        string sColour
    utBorder Border
      [0]
        num nBorderWidth
        string sBorderColour
        string sBorderStyle
    utCommon Common
      [0]
        string sID = "lbl_Title"
        string sPage = "Disk://SmartTCP_CS9/ts2/interface/Page_Main"
        string sText = "史陶比尔工具标定 - SmartTCP"
    utData Data
      [0]
        bool bStatus
        num nVal = 99
    utEvents Events
      [0]
        bool bClick
        bool bMouseDown
        bool bMouseUp
    utText Text
      [0]
        num nFontSize
        string sFontFamily
        string sFontStyle
        string sFontWeight
        string sTextAlignment
public utLabel utLbl_Tool
  [0]
    utAppearance Appearance
      [0]
        bool bVisibility
        string sBackgroundColour = "#FFFFFF"
        string sColour
    utBorder Border
      [0]
        num nBorderWidth
        string sBorderColour
        string sBorderStyle
    utCommon Common
      [0]
        string sID = "lbl_Tool"
        string sPage = "Disk://SmartTCP_CS9/ts2/interface/Page_Main"
        string sText = "工具："
    utData Data
      [0]
        bool bStatus
        num nVal = 99
    utEvents Events
      [0]
        bool bClick
        bool bMouseDown
        bool bMouseUp
    utText Text
      [0]
        num nFontSize
        string sFontFamily
        string sFontStyle
        string sFontWeight
        string sTextAlignment
public utLabel utLbl_ToolValue_Data[6]
  [0]
    utAppearance Appearance
      [0]
        bool bVisibility
        string sBackgroundColour = "#FFFFFF"
        string sColour
    utBorder Border
      [0]
        num nBorderWidth
        string sBorderColour
        string sBorderStyle
    utCommon Common
      [0]
        string sID = "utLbl_ToolValue_Data0"
        string sPage = "Disk://SmartTCP_CS9/ts2/interface/Page_Container_Test"
        string sText = "120    "
    utData Data
      [0]
        bool bStatus
        num nVal = 99
    utEvents Events
      [0]
        bool bClick
        bool bMouseDown
        bool bMouseUp
    utText Text
      [0]
        num nFontSize
        string sFontFamily
        string sFontStyle
        string sFontWeight
        string sTextAlignment
  [1]
    utAppearance Appearance
      [0]
        bool bVisibility
        string sBackgroundColour = "#FFFFFF"
        string sColour
    utBorder Border
      [0]
        num nBorderWidth
        string sBorderColour
        string sBorderStyle
    utCommon Common
      [0]
        string sID = "utLbl_ToolValue_Data1"
        string sPage = "Disk://SmartTCP_CS9/ts2/interface/Page_Container_Test"
        string sText = "55    "
    utData Data
      [0]
        bool bStatus
        num nVal = 99
    utEvents Events
      [0]
        bool bClick
        bool bMouseDown
        bool bMouseUp
    utText Text
      [0]
        num nFontSize
        string sFontFamily
        string sFontStyle
        string sFontWeight
        string sTextAlignment
  [2]
    utAppearance Appearance
      [0]
        bool bVisibility
        string sBackgroundColour = "#FFFFFF"
        string sColour
    utBorder Border
      [0]
        num nBorderWidth
        string sBorderColour
        string sBorderStyle
    utCommon Common
      [0]
        string sID = "utLbl_ToolValue_Data2"
        string sPage = "Disk://SmartTCP_CS9/ts2/interface/Page_Container_Test"
        string sText = "0    "
    utData Data
      [0]
        bool bStatus
        num nVal = 99
    utEvents Events
      [0]
        bool bClick
        bool bMouseDown
        bool bMouseUp
    utText Text
      [0]
        num nFontSize
        string sFontFamily
        string sFontStyle
        string sFontWeight
        string sTextAlignment
  [3]
    utAppearance Appearance
      [0]
        bool bVisibility
        string sBackgroundColour = "#FFFFFF"
        string sColour
    utBorder Border
      [0]
        num nBorderWidth
        string sBorderColour
        string sBorderStyle
    utCommon Common
      [0]
        string sID = "utLbl_ToolValue_Data3"
        string sPage = "Disk://SmartTCP_CS9/ts2/interface/Page_Container_Test"
        string sText = "0    "
    utData Data
      [0]
        bool bStatus
        num nVal = 99
    utEvents Events
      [0]
        bool bClick
        bool bMouseDown
        bool bMouseUp
    utText Text
      [0]
        num nFontSize
        string sFontFamily
        string sFontStyle
        string sFontWeight
        string sTextAlignment
  [4]
    utAppearance Appearance
      [0]
        bool bVisibility
        string sBackgroundColour = "#FFFFFF"
        string sColour
    utBorder Border
      [0]
        num nBorderWidth
        string sBorderColour
        string sBorderStyle
    utCommon Common
      [0]
        string sID = "utLbl_ToolValue_Data4"
        string sPage = "Disk://SmartTCP_CS9/ts2/interface/Page_Container_Test"
        string sText = "0    "
    utData Data
      [0]
        bool bStatus
        num nVal = 99
    utEvents Events
      [0]
        bool bClick
        bool bMouseDown
        bool bMouseUp
    utText Text
      [0]
        num nFontSize
        string sFontFamily
        string sFontStyle
        string sFontWeight
        string sTextAlignment
  [5]
    utAppearance Appearance
      [0]
        bool bVisibility
        string sBackgroundColour = "#FFFFFF"
        string sColour
    utBorder Border
      [0]
        num nBorderWidth
        string sBorderColour
        string sBorderStyle
    utCommon Common
      [0]
        string sID = "utLbl_ToolValue_Data5"
        string sPage = "Disk://SmartTCP_CS9/ts2/interface/Page_Container_Test"
        string sText = "0    "
    utData Data
      [0]
        bool bStatus
        num nVal = 99
    utEvents Events
      [0]
        bool bClick
        bool bMouseDown
        bool bMouseUp
    utText Text
      [0]
        num nFontSize
        string sFontFamily
        string sFontStyle
        string sFontWeight
        string sTextAlignment
public utLabel utLbl_Tool_Data
  [0]
    utAppearance Appearance
      [0]
        bool bVisibility
        string sBackgroundColour = "#FFFFFF"
        string sColour
    utBorder Border
      [0]
        num nBorderWidth
        string sBorderColour
        string sBorderStyle
    utCommon Common
      [0]
        string sID = "lbl_Tool_Data"
        string sPage = "Disk://SmartTCP_CS9/ts2/interface/Page_Main"
        string sText = "tFlange"
    utData Data
      [0]
        bool bStatus
        num nVal = 99
    utEvents Events
      [0]
        bool bClick
        bool bMouseDown
        bool bMouseUp
    utText Text
      [0]
        num nFontSize
        string sFontFamily
        string sFontStyle
        string sFontWeight
        string sTextAlignment
public utText utTxt_OffsetValue_Data[6]
  [0]
    utAppearance Appearance
      [0]
        bool bVisibility
        string sBackgroundColour = "#EEFF00"
        string sColour
    utBorder Border
      [0]
        string sBorderColour
        string sBorderSytle
        string sBorderWidth
    utCommon Common
      [0]
        bool bDisabled
        num nValue
        string sID = "utTxt_OffsetValue_Data0"
        string sPage = "Disk://SmartTCP_CS9/ts2/interface/Page_Container_Test"
        string sValue
    utText Text
      [0]
        num nFontSize
        string sFontFamily
        string sFontStyle
        string sFontWeight
        string sTextAlignment
  [1]
    utAppearance Appearance
      [0]
        bool bVisibility
        string sBackgroundColour = "#EEFF00"
        string sColour
    utBorder Border
      [0]
        string sBorderColour
        string sBorderSytle
        string sBorderWidth
    utCommon Common
      [0]
        bool bDisabled
        num nValue
        string sID = "utTxt_OffsetValue_Data1"
        string sPage = "Disk://SmartTCP_CS9/ts2/interface/Page_Container_Test"
        string sValue
    utText Text
      [0]
        num nFontSize
        string sFontFamily
        string sFontStyle
        string sFontWeight
        string sTextAlignment
  [2]
    utAppearance Appearance
      [0]
        bool bVisibility
        string sBackgroundColour = "#EEFF00"
        string sColour
    utBorder Border
      [0]
        string sBorderColour
        string sBorderSytle
        string sBorderWidth
    utCommon Common
      [0]
        bool bDisabled
        num nValue = 10
        string sID = "utTxt_OffsetValue_Data2"
        string sPage = "Disk://SmartTCP_CS9/ts2/interface/Page_Container_Test"
        string sValue
    utText Text
      [0]
        num nFontSize
        string sFontFamily
        string sFontStyle
        string sFontWeight
        string sTextAlignment
  [3]
    utAppearance Appearance
      [0]
        bool bVisibility
        string sBackgroundColour = "#EEFF00"
        string sColour
    utBorder Border
      [0]
        string sBorderColour
        string sBorderSytle
        string sBorderWidth
    utCommon Common
      [0]
        bool bDisabled
        num nValue
        string sID = "utTxt_OffsetValue_Data3"
        string sPage = "Disk://SmartTCP_CS9/ts2/interface/Page_Container_Test"
        string sValue
    utText Text
      [0]
        num nFontSize
        string sFontFamily
        string sFontStyle
        string sFontWeight
        string sTextAlignment
  [4]
    utAppearance Appearance
      [0]
        bool bVisibility
        string sBackgroundColour = "#EEFF00"
        string sColour
    utBorder Border
      [0]
        string sBorderColour
        string sBorderSytle
        string sBorderWidth
    utCommon Common
      [0]
        bool bDisabled
        num nValue
        string sID = "utTxt_OffsetValue_Data4"
        string sPage = "Disk://SmartTCP_CS9/ts2/interface/Page_Container_Test"
        string sValue
    utText Text
      [0]
        num nFontSize
        string sFontFamily
        string sFontStyle
        string sFontWeight
        string sTextAlignment
  [5]
    utAppearance Appearance
      [0]
        bool bVisibility
        string sBackgroundColour = "#EEFF00"
        string sColour
    utBorder Border
      [0]
        string sBorderColour
        string sBorderSytle
        string sBorderWidth
    utCommon Common
      [0]
        bool bDisabled
        num nValue
        string sID = "utTxt_OffsetValue_Data5"
        string sPage = "Disk://SmartTCP_CS9/ts2/interface/Page_Container_Test"
        string sValue
    utText Text
      [0]
        num nFontSize
        string sFontFamily
        string sFontStyle
        string sFontWeight
        string sTextAlignment
public utText utTxt_popUpMsg
  [0]
    utAppearance Appearance
      [0]
        bool bVisibility
        string sBackgroundColour = "#7C95FF"
        string sColour
    utBorder Border
      [0]
        string sBorderColour
        string sBorderSytle
        string sBorderWidth
    utCommon Common
      [0]
        bool bDisabled
        num nValue
        string sID = "txt_popUpMsg"
        string sPage = "Disk://SmartTCP_CS9/ts2/interface/Page_Container_Confirm"
        string sValue = "第2点记录完成"
    utText Text
      [0]
        num nFontSize
        string sFontFamily
        string sFontStyle
        string sFontWeight
        string sTextAlignment
public utTool utCurrentTool
  [0]
    num nItem
    num nItemM = 1
    string sName
    tool tValue = {fatherId=flange[0]}

--- changeBckColorLabel.pgx ---
public program changeBckColorLabel(utLabel x_uUtLabel, string x_sColor)
begin
  // change the BackGround color -> using userPageSet
  userPageSet(x_uUtLabel.Common.sPage,x_uUtLabel.Common.sID,"style.backgroundColor",x_sColor)
end

--- CheckPosEqual.pgx ---
program CheckPosEqual(point x_pA, bool& x_bPos)
  local point l_pHere
begin
  l_pHere=here(utCurrentTool.tValue,world)
  if power(x_pA.trsf.x-l_pHere.trsf.x,2)+power(x_pA.trsf.y-l_pHere.trsf.y,2)+power(x_pA.trsf.z-l_pHere.trsf.z,2)+power(x_pA.trsf.rz-l_pHere.trsf.rz,2)<0.2
    x_bPos=true
  else
    x_bPos=false
  endIf
//  if power(x_pA.trsf.x-l_pHere.trsf.x,2)+power(x_pA.trsf.y-l_pHere.trsf.y,2)+power(x_pA.trsf.z-l_pHere.trsf.z,2)+power(x_pA.trsf.rx-l_pHere.trsf.rx,2)+power(x_pA.trsf.ry-l_pHere.trsf.ry,2)+power(x_pA.trsf.rz-l_pHere.trsf.rz,2)<1
//    x_bPos=true
//  else
//    x_bPos=false
//  endIf
end

--- CheckTraj.pgx ---
program CheckTraj(point x_pStart, trsf x_trOffset, point x_pEnd, bool& x_bTrajOK)
  local bool l_bOk
  local bool l_bOut
  local num l_nStep
  local trsf l_trMiniOffset
  local trsf l_trStepOffset
  local num l_nVal
  local point l_pTarget
  local jointRs l_jNearBy
  local jointRs l_jTarget
  local jointRs l_jStart
  local point l_pNearBy
  local string l_sPopMsg
begin
  l_trMiniOffset={x_trOffset.x/1000,x_trOffset.y/1000,x_trOffset.z/1000,x_trOffset.rx/1000,x_trOffset.ry/1000,x_trOffset.rz/1000}
  x_pEnd=appro(x_pStart,x_trOffset)
  l_nStep=0
  l_nVal=1
  do
    switch l_nStep
      //******************************************************************
      //Check NearBy Position
      case 0
        l_bOk=pointToJoint(utCurrentTool.tValue,herej(),x_pStart,l_jStart)
        if l_bOk==true
          l_nStep=1
        else
          l_nStep=99
        endIf
      break
      //
      case 1
        l_pNearBy=appro(x_pStart,l_trMiniOffset)
        l_bOk=pointToJoint(utCurrentTool.tValue,herej(),l_pNearBy,l_jNearBy)
        if l_bOk==true
          l_nStep=2
        else
          l_nStep=99
        endIf
      break
      //******************************************************************
      //******************************************************************
      case 2
        l_trStepOffset={x_trOffset.x*l_nVal/100,x_trOffset.y*l_nVal/100,x_trOffset.z*l_nVal/100,x_trOffset.rx*l_nVal/100,x_trOffset.ry*l_nVal/100,x_trOffset.rz*l_nVal/100}
        l_pTarget=appro(x_pStart,l_trStepOffset)
        l_bOk=pointToJoint(utCurrentTool.tValue,herej(),l_pTarget,l_jTarget)
        if l_bOk==true
          l_nStep=3
        else
          l_nStep=99
        endIf
      break
      //
      case 3
        if l_jNearBy.j4-l_jStart.j4>=0 and l_jTarget.j4-l_jStart.j4<0
          l_jTarget.j4=l_jTarget.j4+360
        endIf
        if l_jNearBy.j4-l_jStart.j4<0 and l_jTarget.j4-l_jStart.j4>=0
          l_jTarget.j4=l_jTarget.j4-360
        endIf
        l_nStep=4
      break
      //
      case 4
        if isInRange(l_jTarget)==true
          l_nStep=5
        else
          l_nStep=99
        endIf
      break
      //
      case 5
        if l_nVal<100
          l_nVal=l_nVal+1
          l_nStep=2
        else
          l_nStep=100
        endIf
      break
      //******************************************************************
      case 99
        call updateStr(121,l_sPopMsg,"The maximum rotation angle is only:")
        l_nVal=l_nVal-1
        l_sPopMsg=l_sPopMsg+toString(".",roundDown(l_nVal))+"°"
        popUpMsg(l_sPopMsg)
        //
        x_bTrajOK=false
        l_bOut=true
      break
      case 100
        x_bTrajOK=true
        l_bOut=true
      break
    endSwitch
  until l_bOut
end

--- hmiAlert.pgx ---
public program hmiAlert(string x_sMsg, string x_sMsgType)
  local string l_sMsg
begin
  switch sLanguage
    case "english"
      l_sMsg=sAlertEN[x_sMsg]
    break
    case "chinese"
      l_sMsg=sAlertCN[x_sMsg]
    break
  endSwitch
  //*************************************************************
  utCtn_Message.Common.sSource="Page_Container_Alert.html"
  utTxt_popUpMsg.Common.sValue=l_sMsg
  //*************************************************************
  switch x_sMsgType
    case "info"
      utTxt_popUpMsg.Appearance.sBackgroundColour="#7C95FF"
    break
    //
    case "warning"
      utTxt_popUpMsg.Appearance.sBackgroundColour="#EEFB45"
    break
    //
    case "confirm"
      utTxt_popUpMsg.Appearance.sBackgroundColour="#FFFFFF"
    break
    //
    default
      utTxt_popUpMsg.Appearance.sBackgroundColour="#ADADB2"
    break
  endSwitch
  //*************************************************************
  if taskStatus("HmiClose")!=-1
    taskKill("HmiClose")
  endIf
  if taskStatus("HmiClose")==-1
    taskCreate "HmiClose",100,hmiClose()
  endIf
end

--- hmiClose.pgx ---
public program hmiClose()
  local bool l_bOut
begin
  delay(0.2)
  utCtn_Message.Appearance.bVisibility=true
  //
  l_bOut=false
  nClock=clock()
  do
    if utCtn_Message.Appearance.bVisibility==true
      if clock()-nClock>=3
        utTxt_popUpMsg.Common.sValue=""
        utCtn_Message.Appearance.bVisibility=false
        l_bOut=true
      endIf
      if utBtn_OK.Events.bClick==true
        utBtn_OK.Events.bClick=false
        utTxt_popUpMsg.Common.sValue=""
        utCtn_Message.Appearance.bVisibility=false
        l_bOut=true
      endIf
    endIf
    delay(0)
  until l_bOut
end

--- hmiConfirm.pgx ---
public program hmiConfirm(string x_sMsg, string x_sMsgType, bool& x_bOK)
  local string l_sMsg
  local bool l_bOut
begin
  switch sLanguage
    case "english"
      l_sMsg=sAlertEN[x_sMsg]
    break
    case "chinese"
      l_sMsg=sAlertCN[x_sMsg]
    break
  endSwitch
  //*************************************************************
  utCtn_Message.Common.sSource="Page_Container_Confirm.html"
  utTxt_popUpMsg.Common.sValue=l_sMsg
  //*************************************************************
  switch x_sMsgType
    case "info"
      utTxt_popUpMsg.Appearance.sBackgroundColour="#7C95FF"
    break
    //
    case "warning"
      utTxt_popUpMsg.Appearance.sBackgroundColour="#EEFB45"
    break
    //
    case "confirm"
      utTxt_popUpMsg.Appearance.sBackgroundColour="#FFFFFF"
    break
    //
    default
      utTxt_popUpMsg.Appearance.sBackgroundColour="#ADADB2"
    break
  endSwitch
  delay(0.2)
  //
  utCtn_Message.Appearance.bVisibility=true
  //
  utBtn_Yes.Events.bClick=false
  utBtn_No.Events.bClick=false
  l_bOut=false
  do
    if utBtn_Yes.Events.bClick==true
      utBtn_Yes.Events.bClick=false
      l_bOut=true
      x_bOK=true
    elseIf utBtn_No.Events.bClick==true
      utBtn_No.Events.bClick=false
      l_bOut=true
      x_bOK=false
    endIf
  until l_bOut
  delay(0)
  utCtn_Message.Appearance.bVisibility=false
end

--- initButton.pgx ---
public program initButton(utButton& x_utButton[], string x_sPage, string x_sId, string x_sText)
begin
  x_utButton.Common.sPage=x_sPage
  x_utButton.Common.sID=x_sId
  x_utButton.Common.sText=x_sText
  //
  //userPageBind(x_sPage,x_utButton.Common.sID,"style.backgroundColor",x_utButton.Appearance.sBackgroundColour,1,"r")
  userPageBind(x_utButton.Common.sPage,x_utButton.Common.sID,"innerHTML",x_utButton.Common.sText,1,"r")
  userPageBind(x_utButton.Common.sPage,x_utButton.Common.sID,"style.visibility",x_utButton.Appearance.bVisibility,1,"r")
  userPageBindClick(x_utButton.Common.sPage,x_utButton.Common.sID,x_utButton.Events.bClick,true)
  //
  x_utButton.Appearance.bVisibility=(x_sText!="")
  x_utButton.Events.bClick=false
end

--- initCheckBox.pgx ---
public program initCheckBox(utImage& x_utImage[], string x_sPage, string x_sId, string x_sSatus)
begin
  x_utImage.Common.sPage=x_sPage
  x_utImage.Common.sID=x_sId
  switch x_sSatus
    case "CheckOn"
      x_utImage.Data.sSourceImg1="images/checkbox_checked.png"
      x_utImage.Data.sSourceImg2="images/checkbox_unchecked.png"
      x_utImage.Common.sSourceImage=x_utImage.Data.sSourceImg1
      x_utImage.Data.bStatus=true
    break
    case "CheckOff"
      x_utImage.Data.sSourceImg1="images/checkbox_checked.png"
      x_utImage.Data.sSourceImg2="images/checkbox_unchecked.png"
      x_utImage.Common.sSourceImage=x_utImage.Data.sSourceImg2
      x_utImage.Data.bStatus=false
    break
    case "SwitchOn"
      x_utImage.Data.sSourceImg1="images/switch_on.png"
      x_utImage.Data.sSourceImg2="images/switch_off.png"
      x_utImage.Common.sSourceImage=x_utImage.Data.sSourceImg1
      x_utImage.Data.bStatus=true
    break
    case "SwitchOff"
      x_utImage.Data.sSourceImg1="images/switch_on.png"
      x_utImage.Data.sSourceImg2="images/switch_off.png"
      x_utImage.Common.sSourceImage=x_utImage.Data.sSourceImg2
      x_utImage.Data.bStatus=false
    break
  endSwitch
  //
  userPageBind(x_utImage.Common.sPage,x_utImage.Common.sID,"src",x_utImage.Common.sSourceImage,1,"r")
  userPageBind(x_utImage.Common.sPage,x_utImage.Common.sID,"className",x_utImage.Common.sClass,1,"r")
  userPageBindClick(x_utImage.Common.sPage,x_utImage.Common.sID,x_utImage.Events.bClick,true)
  x_utImage.Events.bClick=false
  x_utImage.Common.sClass="clickable"
end

--- initCombo.pgx ---
public program initCombo(utCombo& x_utCombo[], string x_sPage, string x_sId)
begin
  x_utCombo.Common.sPage=x_sPage
  x_utCombo.Common.sID=x_sId
  userPageBind(x_utCombo.Common.sPage,x_utCombo.Common.sID,"options",x_utCombo.Common.sItem,size(x_utCombo.Common.sItem),"r")
  userPageBind(x_utCombo.Common.sPage,x_utCombo.Common.sID,"value",x_utCombo.Common.sValue,1,"rw")
end

--- initContainer.pgx ---
public program initContainer(utContainer& x_utContainer[], string x_sPage, string x_sId, bool x_bVisibility)
begin
  x_utContainer.Common.sPage=x_sPage
  x_utContainer.Common.sID=x_sId
  userPageBind(x_utContainer.Common.sPage,x_utContainer.Common.sID,"src",x_utContainer.Common.sSource,1,"r")
  userPageBind(x_utContainer.Common.sPage,x_utContainer.Common.sID,"style.visibility",x_utContainer.Appearance.bVisibility,1,"r")
  //
  x_utContainer.Appearance.bVisibility=x_bVisibility
end

--- initImage.pgx ---
public program initImage(utImage& x_utImage[], string x_sPage, string x_sId)
begin
  x_utImage.Common.sPage=x_sPage
  x_utImage.Common.sID=x_sId
  userPageBind(x_utImage.Common.sPage,x_utImage.Common.sID,"src",x_utImage.Common.sSourceImage,1,"r")
  userPageBind(x_utImage.Common.sPage,x_utImage.Common.sID,"style.visibility",x_utImage.Appearance.bVisibility,1,"r")
  userPageBindClick(x_utImage.Common.sPage,x_utImage.Common.sID,x_utImage.Events.bClick,true)
  //
  userPageBind(x_utImage.Common.sPage,x_utImage.Common.sID,"className",x_utImage.Common.sClass,1,"r")
  //userPageBind(x_sPage,x_utImage.Common.sID,"style.borderColor",x_utImage.Border.sBorderColour,1,"r")
  //userPageBind(x_sPage,x_utImage.Common.sID,"style.borderStyle",x_utImage.Border.sBorderStyle,1,"r")
  //
  x_utImage.Appearance.bVisibility=true
  x_utImage.Events.bClick=false
  x_utImage.Common.sClass="clickable"
end

--- initLabel.pgx ---
public program initLabel(utLabel& x_utLabel[], string x_sPage, string x_sId, string x_sText)
begin
  x_utLabel.Common.sPage=x_sPage
  x_utLabel.Common.sID=x_sId
  userPageBind(x_utLabel.Common.sPage,x_utLabel.Common.sID,"innerHTML",x_utLabel.Common.sText,1,"r")
  //userPageBind(x_sPage,x_utLabel.Common.sID,"style.backgroundColor",x_utLabel.Appearance.sBackgroundColour,1,"r")
  //userPageBindClick(x_sPage,x_utLabel.Common.sID,x_utLabel.Events.bClick,true)
  //
  if x_sText=="" or x_sText=="Null"
    x_utLabel.Common.sText=""
  else
    x_utLabel.Common.sText=x_sText
  endIf
  //x_utLabel.Appearance.sBackgroundColour="#F3F4F4"
  x_utLabel.Data.nVal=99
end

--- initList.pgx ---
public program initList(utList& x_utList[], string x_sPage, string x_sId)
begin
  x_utList.Common.sPage=x_sPage
  x_utList.Common.sID=x_sId
  userPageBind(x_utList.Common.sPage,x_utList.Common.sID,"options",x_utList.Common.sItem,size(x_utList.Common.sItem),"r")
  userPageBind(x_utList.Common.sPage,x_utList.Common.sID,"value",x_utList.Common.sValue,1,"rw")
end

--- initText.pgx ---
public program initText(utText& x_utText, string x_sPage, string x_sId, string x_sType)
begin
  x_utText.Common.sPage=x_sPage
  x_utText.Common.sID=x_sId
  switch x_sType
    case "Num"
      userPageBind(x_utText.Common.sPage,x_utText.Common.sID,"value",x_utText.Common.nValue,1,"rw")
    break
    case "String"
      userPageBind(x_utText.Common.sPage,x_utText.Common.sID,"value",x_utText.Common.sValue,1,"rw")
    break
  endSwitch
  userPageBind(x_utText.Common.sPage,x_utText.Common.sID,"style.backgroundColor",x_utText.Appearance.sBackgroundColour,1,"r")
  //
  x_utText.Appearance.sBackgroundColour="trasparent"
  //
end

--- ListMove.pgx ---
public program ListMove(string x_sM)
  local bool l_bA
  local bool l_bB
  local bool l_bC
  local bool l_bEqual
  local frame l_fFrame
  local trsf l_trA
  local point l_pCurrentPosUp
  local point l_pTargetPosUp
  local num l_nJogMode
  local joint l_jTargetPosUp
  local bool l_bOut
  local num l_nStep
  local joint l_jStart
  local point l_pTraj
  local jointRs l_jPos
  local joint l_jCurrentPosUp
  local trsf l_trB
  local pointRs l_pB
  local pointRs l_pA
begin
  resetMotion()
  link(l_pCurrentPosUp,world)
  link(l_pTargetPosUp,world)
  //
  l_nJogMode=nJogMode
  $jogMode(0)
  wait($getJogmode()==0)
  delay(0.1)
  //
  //*******************************************************************************************
  switch x_sM
    case "pTeach1"
    call moveTarget(pTeach1,jTeach1)
    break
    //
    case "pTeach2"
    call moveTarget(pTeach2,jTeach2)
    break
    //
    case "pTeach3"
     call moveTarget(pTeach3,jTeach3)
    break
    //
    case "pTeach4"
     call moveTarget(pTeach4,jTeach4)
    break
    //
    case "pTeach5"
      call moveTarget(pTeach5,jTeach5)
    break
    //
    case "pTeach6"
      call moveTarget(pTeach6,jTeach6)
    break
    //*******************************************************************************************
    case "pAdjustXY_2_1"
      call moveTarget(pAdjustXY_2_1,jAdjustXY_2_1)
    break
    //
    case "pAdjustXY_2_2"
      call moveTarget(pAdjustXY_2_2,jAdjustXY_2_2)
    break
    //
    case "pAdjustXY_3_1"
      call moveTarget(pAdjustXY_3_1,jAdjustXY_3_1)
    break
    //
    case "pAdjustXY_3_2"
      call moveTarget(pAdjustXY_3_2,jAdjustXY_3_2)
    break
    //
    case "pAdjustXY_3_3"
      call moveTarget(pAdjustXY_3_3,jAdjustXY_3_3)
    break
    //*******************************************************************************************
  case "GoBack_pAdjustXY_2_1"
      l_bOut=false
      l_nStep=0
      do
        switch l_nStep
          case 0
            if pAdjustXY_2_1.trsf!={0,0,0,0,0,0}
              l_nStep=1
            else
              l_nStep=99
            endIf
          break
          //
          case 1
            call CheckPosEqual(pAdjustXY_2_1,l_bEqual)
            if l_bEqual==true
              l_nStep=100
            else
              l_nStep=2
            endIf
          break
          //
          case 2
            call CheckPosEqual(pAdjustXY_2_2,l_bEqual)
            if l_bEqual==true
              l_nStep=3
            else
              l_nStep=4
            endIf
          break
          //
          case 3
              call hmiAlert("GoBack","info")
              movel(_pA,utCurrentTool.tValue,mSpeed_C_blend)
              movel(pAdjustXY_2_1,utCurrentTool.tValue,mSpeed_C_blend)
              waitEndMove()
              l_nStep=100
          break
          //
          case 4
            l_pCurrentPosUp=compose(here(utCurrentTool.tValue,world),world,{0,0,20,0,0,0})
            l_pTargetPosUp=appro(pAdjustXY_2_1,{0,0,-20,0,0,0})
            l_bA=pointToJoint(utCurrentTool.tValue,jAdjustXY_2_1,l_pTargetPosUp,l_jTargetPosUp)
            if l_bA==true
              call hmiAlert("GoBack","info")
              movel(l_pCurrentPosUp,utCurrentTool.tValue,mSpeed_J_blend)
              movej(l_jTargetPosUp,utCurrentTool.tValue,mSpeed_J_blend)
              movel(pAdjustXY_2_1,utCurrentTool.tValue,mSlow)
              waitEndMove()
              l_nStep=100
            else
              l_nStep=99
            endIf
          break
          //
          case 99
            call hmiAlert("CantGoBack","warning")
            l_bOut=true
          break
          //
          case 100
            call hmiAlert("CompleteGoBack","info")
            l_bOut=true
          break
        endSwitch
      until l_bOut
    break
    //
    case "Rz+180_pAdjustXY_2_1"
      l_bOut=false
      l_nStep=0
      do
        switch l_nStep
          case 0
            l_trA={0,0,0,0,0,90}
            l_trB={0,0,0,0,0,180}
            l_pA=appro(pAdjustXY_2_1,l_trA)
            l_pB=appro(pAdjustXY_2_1,l_trB)
            l_pA.config=cConfigSame
            l_pB.config=cConfigSame
            //
            call CheckPosEqual(l_pB,l_bEqual)
            if l_bEqual==true
              l_nStep=100
            else
              call CheckTraj(pAdjustXY_2_1,l_trA,l_pA,l_bA)
              call CheckTraj(pAdjustXY_2_1,l_trB,l_pB,l_bB)
              l_nStep=1
            endIf
          break
          //
          case 1
            //whether the target position is reachable
            if l_bA==true and l_bB==true
              l_nStep=2
            else
              l_nStep=99
            endIf
          break
          //
          case 2
            //Whether the robot is at the end position
            call CheckPosEqual(l_pB,l_bEqual)
            if !l_bEqual
              l_nStep=3
            else
              l_nStep=100
            endIf
          break
          //
          case 3
            call hmiAlert("Move","info")
            _pA=l_pA
            _pB=l_pB
            movel(_pA,utCurrentTool.tValue,mSpeed_C_blend)
            movel(_pB,utCurrentTool.tValue,mSpeed_C_blend)
            waitEndMove()
            l_nStep=100
          break
          //
          case 99
            call hmiAlert("CantMove1","warning")
            l_bOut=true
          break
          //
          case 100
            call hmiAlert("CompleteMove","info")
            l_bOut=true
          break
        endSwitch
      until l_bOut
    break
    //
    case "Rz-180_pAdjustXY_2_1"
      l_bOut=false
      l_nStep=0
      do
        switch l_nStep
          case 0
            l_trA={0,0,0,0,0,-90}
            l_trB={0,0,0,0,0,-180}
            l_pA=appro(pAdjustXY_2_1,l_trA)
            l_pB=appro(pAdjustXY_2_1,l_trB)
            l_pA.config=cConfigSame
            l_pB.config=cConfigSame
            //
            call CheckPosEqual(l_pB,l_bEqual)
            if l_bEqual==true
              l_nStep=100
            else
              call CheckTraj(pAdjustXY_2_1,l_trA,l_pA,l_bA)
              call CheckTraj(pAdjustXY_2_1,l_trB,l_pB,l_bB)
              l_nStep=1
            endIf
          break
          //
          case 1
            //whether the target position is reachable
            if l_bA==true and l_bB==true
              l_nStep=2
            else
              l_nStep=99
            endIf
          break
          //
          case 2
            //Whether the robot is at the end position
            call CheckPosEqual(l_pB,l_bEqual)
            if !l_bEqual
              l_nStep=3
            else
              l_nStep=100
            endIf
          break
          //
          case 3
            call hmiAlert("Move","info")
            _pA=l_pA
            _pB=l_pB
            movel(_pA,utCurrentTool.tValue,mSpeed_C_blend)
            movel(_pB,utCurrentTool.tValue,mSpeed_C_blend)
            waitEndMove()
            l_nStep=100
          break
          //
          case 99
            call hmiAlert("CantMove1","warning")
            l_bOut=true
          break
          //
          case 100
            call hmiAlert("CompleteMove","info")
            l_bOut=true
          break
        endSwitch
      until l_bOut
    break
    //
    case "GoBack_pAdjustXY_3_1"
      if pAdjustXY_3_1.trsf!={0,0,0,0,0,0}
        call CheckPosEqual(pAdjustXY_3_1,l_bEqual)
        if l_bEqual
          //At the starting positio
          call hmiAlert("CompleteGoBack","info")
        else
          //Not At the starting position
          call hmiAlert("GoBack","info")
          movel(pAdjustXY_3_1,utCurrentTool.tValue,mSpeed_C_blend)
          waitEndMove()
          call hmiAlert("CompleteGoBack","info")
        endIf
      else
        call hmiAlert("CantGoBack","warning")
      endIf
    break
    //
    case "Rz+60_pAdjustXY_3_1"
      l_bOut=false
      l_nStep=0
      do
        switch l_nStep
          case 0
            l_trA={0,0,0,0,0,60}
            _pA=appro(pAdjustXY_3_1,l_trA)
            _pA.config=cConfigSame
            //
            call CheckPosEqual(_pA,l_bEqual)
            if l_bEqual==true
              l_nStep=100
            else
              call CheckTraj(pAdjustXY_3_1,l_trA,_pA,l_bA)
              l_nStep=1
            endIf
          break
          //
          case 1
            //whether the target position is reachable
            if l_bA==true
              l_nStep=2
            else
              l_nStep=99
            endIf
          break
          //
          case 2
            //Whether the robot is at the end position
            call CheckPosEqual(_pA,l_bEqual)
            if !l_bEqual
              l_nStep=3
            else
              l_nStep=100
            endIf
          break
          //
          case 3
            call hmiAlert("Move","info")
            movel(_pA,utCurrentTool.tValue,mSpeed_C_blend)
            waitEndMove()
            l_nStep=100
          break
          //
          case 99
            call hmiAlert("CantMove1","warning")
            l_bOut=true
          break
          //
          case 100
            call hmiAlert("CompleteMove","info")
            l_bOut=true
          break
        endSwitch
      until l_bOut
    break
    //
    case "Rz-60_pAdjustXY_3_1"
      l_bOut=false
      l_nStep=0
      do
        switch l_nStep
          case 0
            l_trA={0,0,0,0,0,-60}
            _pA=appro(pAdjustXY_3_1,l_trA)
            _pA.config=cConfigSame
            //
            call CheckPosEqual(_pA,l_bEqual)
            if l_bEqual==true
              l_nStep=100
            else
              call CheckTraj(pAdjustXY_3_1,l_trA,_pA,l_bA)
              l_nStep=1
            endIf
          break
          //
          case 1
            //whether the target position is reachable
            if l_bA==true
              l_nStep=2
            else
              l_nStep=99
            endIf
          break
          //
          case 2
            //Whether the robot is at the end position
            call CheckPosEqual(_pA,l_bEqual)
            if !l_bEqual
              l_nStep=3
            else
              l_nStep=100
            endIf
          break
          //
          case 3
            call hmiAlert("Move","info")
            movel(_pA,utCurrentTool.tValue,mSpeed_C_blend)
            waitEndMove()
            l_nStep=100
          break
          //
          case 99
            call hmiAlert("CantMove1","warning")
            l_bOut=true
          break
          //
          case 100
            call hmiAlert("CompleteMove","info")
            l_bOut=true
          break
        endSwitch
      until l_bOut
    break
  endSwitch
  $jogMode(l_nJogMode)
end

--- moveTarget.pgx ---
public program moveTarget(point x_pTarget, joint x_jTarget)
  local bool l_bEqual
  local joint l_jCurrentPosUp
  local joint l_jTargetPosUp
  local point l_pCurrentPosUp
  local point l_pTargetPosUp
  local bool l_bOK1
  local bool l_bOK2
begin
  call CheckPosEqual(x_pTarget,l_bEqual)
  if l_bEqual==false
    call hmiAlert("Move","info")
    l_pCurrentPosUp=compose(here(utCurrentTool.tValue,world),world,{0,0,20,0,0,0})
    l_bOK1=pointToJoint(utCurrentTool.tValue,x_jTarget,l_pCurrentPosUp,l_jCurrentPosUp)
    l_pTargetPosUp=appro(x_pTarget,{0,0,-20,0,0,0})
    l_bOK2=pointToJoint(utCurrentTool.tValue,x_jTarget,l_pTargetPosUp,l_jTargetPosUp)
    if l_bOK1==true and l_bOK2==true
      movel(l_pCurrentPosUp,utCurrentTool.tValue,mSpeed_J_blend)
      movej(l_jTargetPosUp,utCurrentTool.tValue,mSpeed_J_blend)
      movel(x_pTarget,utCurrentTool.tValue,mSlow)
      waitEndMove()
      call hmiAlert("CompleteMove","info")
    else
      call hmiAlert("CantMove2","warning")
    endIf
  else
    call hmiAlert("CompleteMove","info")
  endIf
end

--- putMessage.pgx ---
public program putMessage(string x_sMsg, string x_sMsgType)
begin
  switch x_sMsgType
    case "info"
      utTxt_popUpMsg.Appearance.sBackgroundColour="#7C95FF"
    break
    //
    case "warning"
      utTxt_popUpMsg.Appearance.sBackgroundColour="#EEFB45"
    break
    //
    case "confirm"
      utTxt_popUpMsg.Appearance.sBackgroundColour="#FFFFFF"
    break
    //
    default
      utTxt_popUpMsg.Appearance.sBackgroundColour="#ADADB2"
    break
  endSwitch
  utTxt_popUpMsg.Common.sValue=x_sMsg
  delay(0.2)
  utCtn_Message.Appearance.bVisibility=true
end

--- refreshCheckBox.pgx ---
public program refreshCheckBox(utImage& x_utImage[])
  local num l_nI
  local num l_nJ
begin
    if size(x_utImage) != 1
      for l_nI= 0 to size(x_utImage)-1
        if x_utImage[l_nI].Events.bClick==true
          x_utImage[l_nI].Events.bClick=false
          l_nJ=l_nI
          for l_nI=0 to size(x_utImage)-1
            if l_nI==l_nJ
              x_utImage[l_nI].Common.sSourceImage=x_utImage[l_nI].Data.sSourceImg1
              x_utImage[l_nI].Data.bStatus=true
            else
              x_utImage[l_nI].Common.sSourceImage=x_utImage[l_nI].Data.sSourceImg2
              x_utImage[l_nI].Data.bStatus=false
            endIf
          endFor
        endIf
      endFor
    else
      if x_utImage[l_nI].Events.bClick==true
        x_utImage[l_nI].Events.bClick=false
        if x_utImage[l_nI].Data.bStatus==false
          x_utImage[l_nI].Common.sSourceImage=x_utImage[l_nI].Data.sSourceImg1
          x_utImage[l_nI].Data.bStatus=true
        else
          x_utImage[l_nI].Common.sSourceImage=x_utImage[l_nI].Data.sSourceImg2
          x_utImage[l_nI].Data.bStatus=false
        endIf
      endIf
    endIf
end

--- refreshInfo.pgx ---
public program refreshInfo()
begin
  //Version
  if utImg_Info.Events.bClick==true
    utImg_Info.Events.bClick=false
    call hmiAlert("Version","info")
  endIf
end

--- refreshJogMode.pgx ---
public program refreshJogMode()
  local num l_nI
  local pointRs l_pHere
  local jointRs l_jHere
begin
  if workingMode()==1 or workingMode()==2
    for l_nI= 0 to size(utImg_JogMode)-1
      if utImg_JogMode[l_nI].Events.bClick==true
        utImg_JogMode[l_nI].Events.bClick=false
        $jogMode(l_nI)
        nJogMode=$getJogmode()
        switch nJogMode
          case 1
            bShowJpos=true
          break
          case 2,3
            bShowJpos=false
          break
        endSwitch
      endIf
    endFor
  endIf
  //*********************************************************
  if utImg_PosSwitch.Events.bClick==true
    utImg_PosSwitch.Events.bClick=false
    bShowJpos=!bShowJpos
  endIf
  //*********************************************************
  l_pHere=here(utCurrentTool.tValue,world)
  l_jHere=herej()
  if bShowJpos==true
    utLbl_CurrentPos_Name[0].Common.sText="J1:"
    utLbl_CurrentPos_Name[1].Common.sText="J2:"
    utLbl_CurrentPos_Name[2].Common.sText="J3:"
    utLbl_CurrentPos_Name[3].Common.sText="J4:"
    utLbl_CurrentPos_Name[4].Common.sText=""
    utLbl_CurrentPos_Name[5].Common.sText=""
    //
    utLbl_CurrentPos_Data[0].Common.sText=toString(".3",l_jHere.j1)
    utLbl_CurrentPos_Data[1].Common.sText=toString(".3",l_jHere.j2)
    utLbl_CurrentPos_Data[2].Common.sText=toString(".3",l_jHere.j3)
    utLbl_CurrentPos_Data[3].Common.sText=toString(".3",l_jHere.j4)
    utLbl_CurrentPos_Data[4].Common.sText=toString(".3",0)
    utLbl_CurrentPos_Data[5].Common.sText=toString(".3",0)
    //
    utLbl_CurrentPos_Name[4].Appearance.bVisibility=false
    utLbl_CurrentPos_Name[5].Appearance.bVisibility=false
    utLbl_CurrentPos_Data[4].Appearance.bVisibility=false
    utLbl_CurrentPos_Data[5].Appearance.bVisibility=false
  else
    utLbl_CurrentPos_Name[0].Common.sText="X:"
    utLbl_CurrentPos_Name[1].Common.sText="Y:"
    utLbl_CurrentPos_Name[2].Common.sText="Z:"
    utLbl_CurrentPos_Name[3].Common.sText="RX:"
    utLbl_CurrentPos_Name[4].Common.sText="RY:"
    utLbl_CurrentPos_Name[5].Common.sText="RZ:"
    //
    utLbl_CurrentPos_Data[0].Common.sText=toString(".3",l_pHere.trsf.x)
    utLbl_CurrentPos_Data[1].Common.sText=toString(".3",l_pHere.trsf.y)
    utLbl_CurrentPos_Data[2].Common.sText=toString(".3",l_pHere.trsf.z)
    utLbl_CurrentPos_Data[3].Common.sText=toString(".3",l_pHere.trsf.rx)
    utLbl_CurrentPos_Data[4].Common.sText=toString(".3",l_pHere.trsf.ry)
    utLbl_CurrentPos_Data[5].Common.sText=toString(".3",l_pHere.trsf.rz)
    //
    utLbl_CurrentPos_Name[4].Appearance.bVisibility=true
    utLbl_CurrentPos_Name[5].Appearance.bVisibility=true
    utLbl_CurrentPos_Data[4].Appearance.bVisibility=true
    utLbl_CurrentPos_Data[5].Appearance.bVisibility=true
  endIf
  //*********************************************************
  nJogMode=$getJogmode()
  for l_nI= 0 to size(utImg_JogMode)-1
    if l_nI==nJogMode
      //utImg_JogMode[l_nI].Border.sBorderStyle="Solid"
      //utImg_JogMode[l_nI].Border.sBorderColour="#000000"
      utImg_JogMode[l_nI].Common.sClass="selected"
    else
      //utImg_JogMode[l_nI].Border.sBorderStyle="None"
      //utImg_JogMode[l_nI].Border.sBorderColour="#FFFFFF"
      utImg_JogMode[l_nI].Common.sClass="clickable"
    endIf
  endFor
end

--- refreshLanguage.pgx ---
public program refreshLanguage()
begin
  //*************************************************************************************************
  //Get the current robot installation mode
  if sCbxMounting!=utCbx_Mounting_Data.Common.sValue
    sCbxMounting=utCbx_Mounting_Data.Common.sValue
    switch utCbx_Mounting_Data.Common.sValue
      case "置地","Floor"
        sMounting="Floor"
      break
      case "置顶","Ceiling"
        sMounting="Ceiling"
      break
    endSwitch
  endIf

  //*************************************************************************************************
  //Get the current robot interface language
  if sCbxLanguage!=utCbx_Language_Data.Common.sValue
    sCbxLanguage=utCbx_Language_Data.Common.sValue
    switch utCbx_Language_Data.Common.sValue
      case "中文","Chinese"
        sLanguage="chinese"
      break
      //
      case "英文","English"
        sLanguage="english"
      break
      //
      default
        sLanguage="english"
      break
    endSwitch
  endIf
  //*************************************************************************************************
  if sLanguage!=sLanguageM
    sLanguageM=sLanguage
    switch sLanguage
      case "chinese"
        utCbx_Language_Data.Common.sValue="中文"
        utCbx_Language_Data.Common.sItem[0]="中文"
        utCbx_Language_Data.Common.sItem[1]="英文"
        utCbx_Mounting_Data.Common.sItem[0]="置地"
        utCbx_Mounting_Data.Common.sItem[1]="置顶"
        switch utCbx_Mounting_Data.Common.sValue
          case "置地","Floor"
            utCbx_Mounting_Data.Common.sValue="置地"
          break
          case "置顶","Ceiling"
            utCbx_Mounting_Data.Common.sValue="置顶"
          break
        endSwitch
      break
      //
      case "english"
        utCbx_Language_Data.Common.sValue="English"
        utCbx_Language_Data.Common.sItem[0]="English"
        utCbx_Language_Data.Common.sItem[1]="Chinese"
        utCbx_Mounting_Data.Common.sItem[0]="Floor"
        utCbx_Mounting_Data.Common.sItem[1]="Ceiling"
        switch utCbx_Mounting_Data.Common.sValue
          case "置地","Floor"
            utCbx_Mounting_Data.Common.sValue="Floor"
          break
          case "置顶","Ceiling"
            utCbx_Mounting_Data.Common.sValue="Ceiling"
          break
        endSwitch
      break
    endSwitch
    //*************************************************************************************************
        if utBtn_Step[0].Events.bClick==true
      switch nStep0
        case 11,21,31,41,51,61
           nStep0=nStep0-1
        break
       endSwitch
    endIf
    //
    if utBtn_Step[1].Events.bClick==true
      switch nStep1
        case 11,21,31
          nStep1=nStep1-1
        break
      endSwitch
    endIf
    //
    call updateStr(4,utLbl_Title.Common.sText,"Stäubli Tool Calibration - SmartTCP")
    //
    call updateStr(2,utLbl_Language.Common.sText,"Language:")
    //
    call updateStr(3,utLbl_Mounting.Common.sText,"Mounting:")
    //
    call updateStr(7,utLbl_Axis.Common.sText,"ArmType:")
    call updateStr(8,utLbl_Axis_Data.Common.sText,"4axis")
    //
    call updateStr(10,utLbl_Tool.Common.sText,"Tool:")
    //
    call updateStr(11,utLbl_CheckBox_a[0].Common.sText,"2Points")
    call updateStr(12,utLbl_CheckBox_a[1].Common.sText,"3Points")
    call updateStr(13,utLbl_CheckBox_a[2].Common.sText,"6Points")
    //
    call updateStr(14,utLbl_CheckBox_b[0].Common.sText,"2Points180°")
    call updateStr(15,utLbl_CheckBox_b[1].Common.sText,"3Points120°")
    //
    call updateStr(16,utBtn_Step[0].Common.sText,"Calibration tool")
    call updateStr(17,utBtn_Step[1].Common.sText,"Correction tool XY")
    call updateStr(19,utBtn_Step[2].Common.sText,"Verification tool")
    //
    call updateStr(20,utLbl_SwitchTool.Common.sText,"Tool Switch：")
    call updateStr(21,utLbl_Offset.Common.sText,"Tool Offset：")
    //
    call updateStr(utLbl_Point.Data.nVal,utLbl_Point.Common.sText,"")
    call updateStr(utLbl_Step.Data.nVal,utLbl_Step.Common.sText,"")
    //
    call updateInfo(utLbl_Info0.Data.nVal,utLbl_Info0.Data.nVal,utLbl_Info0.Common.sText,"0","")
    call updateInfo(utLbl_Info1.Data.nVal,utLbl_Info1.Data.nVal,utLbl_Info1.Common.sText,"1","")
    call updateInfo(utLbl_Info2.Data.nVal,utLbl_Info2.Data.nVal,utLbl_Info2.Common.sText,"2","")
    call updateInfo(utLbl_Info3.Data.nVal,utLbl_Info3.Data.nVal,utLbl_Info3.Common.sText,"3","")
    call updateInfo(utLbl_Info4.Data.nVal,utLbl_Info4.Data.nVal,utLbl_Info4.Common.sText,"4","")
    //
    call updateBtn(nBtnItem,"Null,Null,Null,Null,Null,Null,Null,Quit")
  endIf
end

--- refreshQuit.pgx ---
public program refreshQuit(bool& x_bOut)
begin
  //Quit
  if utBtn_Step[0].Events.bClick==false and  utBtn_Step[1].Events.bClick==false and utBtn_Step[2].Events.bClick==false
    if utBtn_Bottom[7].Events.bClick==true
      utBtn_Bottom[7].Events.bClick=false
      //Press F7
      call hmiConfirm("Quit","confirm",x_bOut)
    endIf
  endIf
end

--- updateBtn.pgx ---
public program updateBtn(num x_nItemIn, string x_sComment)
  local num l_nI
  local num l_nPos
  local string l_sLongStr
  local string l_sBtnText[8]
begin
  switch sLanguage
    case "chinese"
      l_sLongStr=sHmiCN[x_nItemIn]
    break
    //
    case "english"
      l_sLongStr=sHmiEN[x_nItemIn]
    break
  endSwitch
  nBtnItem=x_nItemIn
  //
  for l_nI= 0 to 7
    l_nPos=find(l_sLongStr,",")
    if l_nPos!=-1
      l_sBtnText[l_nI]=left(l_sLongStr,l_nPos)
      l_sLongStr=delete(l_sLongStr,l_nPos+1,0)
    else
      l_sBtnText[l_nI]=l_sLongStr
    endIf
    if l_sBtnText[l_nI]!="Null"
      utBtn_Bottom[l_nI].Common.sText=l_sBtnText[l_nI]
      utBtn_Bottom[l_nI].Appearance.bVisibility=true
    else
      utBtn_Bottom[l_nI].Common.sText=""
      utBtn_Bottom[l_nI].Appearance.bVisibility=false
    endIf
  endFor
end

--- updateCurrentPos.pgx ---
public program updateCurrentPos()
  local pointRs l_pHere
  local jointRs l_jHere
begin
  nJogMode=$getJogmode()
  switch nJogMode
    case 1
      bShowJpos=true
    break
    case 2,3
      bShowJpos=false
    break
    default
      bShowJpos=true
    break
  endSwitch
  //
  l_pHere=here(utCurrentTool.tValue,world)
  l_jHere=herej()
  if bShowJpos==true
    utLbl_CurrentPos_Name[0].Common.sText="J1:"
    utLbl_CurrentPos_Name[1].Common.sText="J2:"
    utLbl_CurrentPos_Name[2].Common.sText="J3:"
    utLbl_CurrentPos_Name[3].Common.sText="J4:"
    utLbl_CurrentPos_Name[4].Common.sText=""
    utLbl_CurrentPos_Name[5].Common.sText=""
    //
    utLbl_CurrentPos_Data[0].Common.sText=toString(".3",l_jHere.j1)
    utLbl_CurrentPos_Data[1].Common.sText=toString(".3",l_jHere.j2)
    utLbl_CurrentPos_Data[2].Common.sText=toString(".3",l_jHere.j3)
    utLbl_CurrentPos_Data[3].Common.sText=toString(".3",l_jHere.j4)
    utLbl_CurrentPos_Data[4].Common.sText=toString(".3",0)
    utLbl_CurrentPos_Data[5].Common.sText=toString(".3",0)
    //
    utLbl_CurrentPos_Name[4].Appearance.bVisibility=false
    utLbl_CurrentPos_Name[5].Appearance.bVisibility=false
    utLbl_CurrentPos_Data[4].Appearance.bVisibility=false
    utLbl_CurrentPos_Data[5].Appearance.bVisibility=false
  else
    utLbl_CurrentPos_Name[0].Common.sText="X:"
    utLbl_CurrentPos_Name[1].Common.sText="Y:"
    utLbl_CurrentPos_Name[2].Common.sText="Z:"
    utLbl_CurrentPos_Name[3].Common.sText="RX:"
    utLbl_CurrentPos_Name[4].Common.sText="RY:"
    utLbl_CurrentPos_Name[5].Common.sText="RZ:"
    //
    utLbl_CurrentPos_Data[0].Common.sText=toString(".3",l_pHere.trsf.x)
    utLbl_CurrentPos_Data[1].Common.sText=toString(".3",l_pHere.trsf.y)
    utLbl_CurrentPos_Data[2].Common.sText=toString(".3",l_pHere.trsf.z)
    utLbl_CurrentPos_Data[3].Common.sText=toString(".3",l_pHere.trsf.rx)
    utLbl_CurrentPos_Data[4].Common.sText=toString(".3",l_pHere.trsf.ry)
    utLbl_CurrentPos_Data[5].Common.sText=toString(".3",l_pHere.trsf.rz)
    //
    utLbl_CurrentPos_Name[4].Appearance.bVisibility=true
    utLbl_CurrentPos_Name[5].Appearance.bVisibility=true
    utLbl_CurrentPos_Data[4].Appearance.bVisibility=true
    utLbl_CurrentPos_Data[5].Appearance.bVisibility=true
  endIf
end

--- updateInfo.pgx ---
public program updateInfo(num x_nItemIn, num& x_nItemOut, string& x_sTextOut, string x_sNo, string x_sComment)
  local string l_sTextOut
begin
  switch sLanguage
    case "chinese"
      l_sTextOut=sHmiCN[x_nItemIn]
    break
    case "english"
      l_sTextOut=sHmiEN[x_nItemIn]
    break
  endSwitch
  if x_sNo=="0" or x_nItemIn==100
    x_sTextOut=l_sTextOut
  else
    if x_nItemIn==99
      x_sTextOut=""
    else
      x_sTextOut=x_sNo+"."+l_sTextOut
    endIf
  endIf
  x_nItemOut=x_nItemIn
end

--- updateStr.pgx ---
public program updateStr(num x_nItemIn, string& x_sTextOut, string x_sComment)
begin
  switch sLanguage
    case "chinese"
      x_sTextOut=sHmiCN[x_nItemIn]
    break
    //
    case "english"
      x_sTextOut=sHmiEN[x_nItemIn]
    break
  endSwitch
end

--- updateTeachPos.pgx ---
public program updateTeachPos(point x_pteach, bool x_bteach)
begin
  if x_bteach==true
    utLbl_Point.Appearance.sBackgroundColour="#7CFA3F"
  else
    utLbl_Point.Appearance.sBackgroundColour="#FFFFFF"
  endIf
  utLbl_PosValue_Data[0].Common.sText=toString(".3",x_pteach.trsf.x)
  utLbl_PosValue_Data[1].Common.sText=toString(".3",x_pteach.trsf.y)
  utLbl_PosValue_Data[2].Common.sText=toString(".3",x_pteach.trsf.z)
  utLbl_PosValue_Data[3].Common.sText=toString(".3",x_pteach.trsf.rx)
  utLbl_PosValue_Data[4].Common.sText=toString(".3",x_pteach.trsf.ry)
  utLbl_PosValue_Data[5].Common.sText=toString(".3",x_pteach.trsf.rz)
end

--- updateTool.pgx ---
public program updateTool(num x_nToolNumber, bool x_bOffsetActive)
  local bool l_bOut
  local num l_nStep
begin
  l_bOut=false
  l_nStep=0
  do
    switch l_nStep
      case 0
        //Decide which tool to use
        utCurrentTool.nItem=x_nToolNumber
        switch x_nToolNumber
          case 0
            utCurrentTool.tValue=tFlange
            utLbl_Tool_Data.Common.sText="tFlange"
            //call hmiAlert("SwitchFlange")
            l_nStep=1
          break
          case 1
            utCurrentTool.tValue=tTool1
            utLbl_Tool_Data.Common.sText="tTool1"
            //call hmiAlert("SwitchTool1")
            l_nStep=1
          break
          case 2
            utCurrentTool.tValue=tTool2
            utLbl_Tool_Data.Common.sText="tTool2"
            //call hmiAlert("SwitchTool2")
            l_nStep=1
          break
        endSwitch
      break
      //
      case 1
        //Add or not add tool deviations?
        if utImg_Switch.Data.bStatus==true and x_bOffsetActive==true
          utCurrentTool.tValue.trsf=utCurrentTool.tValue.trsf*trOffset
          l_nStep=2
        else
          utCurrentTool.tValue.trsf=utCurrentTool.tValue.trsf
          l_nStep=2
        endIf
      break
      //
      case 2
        //Update current tool value
        tCurrentTool=utCurrentTool.tValue
        $jogContext(tCurrentTool,world,0)
        l_nStep=3
      break
      //
      case 3
        l_bOut=true
      break
    endSwitch
  until l_bOut
end
